Staubli VAL3: refreshInfo.pgx

public program refreshInfo()
begin
  //Version
  if utImg_Info.Events.bClick==true
    utImg_Info.Events.bClick=false
    call hmiAlert("Version","info")
  endIf
end
